Fanuc KAREL source: kd00014.KL

-- PROVISIONAL review KL for V940-1; original PC SHA256 7571825868bb1d49df6b0b348ffc938e83deb8fce81452e3f643251e418b4a7d
-- Incomplete behavior may be omitted. Consult companion uncertainty JSON. Do not deploy.
PROGRAM KD00014
%NOLOCKGROUP
VAR
  I : INTEGER
  J : INTEGER
  B : BOOLEAN
  R : REAL
  S : STRING[80]
BEGIN
  -- V9_ZERO_TABLE_METADATA_HINT layout=0001; no indexed target words; source/name/runtime held
  -- UNRESOLVED_PC offsets 5-9; opcodes 9C,9D,1A
  -- UNRESOLVED_PC offsets 14-18; opcodes 7F
END KD00014
